(* IEC 61131-3 sources: PLC-Static-Analysis/modules/plc-rules/src/test/resources/PLCA-S001, 2 files *)

(* ---- compliant.st ---- *)
TYPE ST_LibVersion :
STRUCT
    iMajor : INT;
    sVersion : STRING;
END_STRUCT
END_TYPE

VAR_GLOBAL
    gstVersion : ST_LibVersion := (iMajor := 1, sVersion := '1.2.0.6');
    gsFirmwareRev : STRING := '3.4.3.0';
END_VAR

FUNCTION_BLOCK FB_ConnOk
VAR_INPUT
    sPassword : STRING;
    sExpected : STRING;
END_VAR
VAR
    sPwd : STRING;
    sHost : STRING;
    sMask : STRING;
    sAms : STRING;
    sMsg : STRING;
    sVersion : STRING;
    nPasswordLength : INT;
    bOk : BOOL;
END_VAR
sPwd := '';
sPassword := '*****';
sHost := '127.0.0.1';
sMask := '255.255.255.0';
sAms := '5.12.34.56.1.1';
sMsg := 'Password wrong';
sVersion := '1.2.3';
sHost := '0.0.0.0';
nPasswordLength := 8;
bOk := sPassword = sExpected;
END_FUNCTION_BLOCK

(* ---- noncompliant.st ---- *)
VAR_GLOBAL
    gsPlcIp : STRING := '10.0.0.15'; // PLCA-S001
    gsApiToken : STRING := 'abc123xyz'; // PLCA-S001
END_VAR

FUNCTION_BLOCK FB_Conn
VAR_INPUT
    sPassword : STRING;
END_VAR
VAR
    sPwd : STRING;
    sHost : STRING;
    bOk : BOOL;
    fbClient : FB_TcpClient;
    wsKennwort : WSTRING := "geheim"; // PLCA-S001
END_VAR
sPwd := 'hunter2'; // PLCA-S001
sHost := '192.168.1.100:502'; // PLCA-S001
bOk := sPassword = 'letmein'; // PLCA-S001
fbClient(sRemoteHost := '172.16.0.2', sPassword := 'admin'); // PLCA-S001 PLCA-S001
END_FUNCTION_BLOCK
